(* IEC 61131-3 sources: tsplc/packages/vscode-extension/tests/fixtures/build-tool/transport/PRG_Transport, 1 file *)

(* ---- declaration.st ---- *)
PROGRAM PRG_Transport
VAR
	Conveyor : FB_Conveyor;
	ClampedSpeed : INT;
END_VAR
